Fanuc KAREL source: KT00657.KL

PROGRAM KT00657
%NOLOCKGROUP
VAR
  P1: POSITION
  P2: POSITION
  OUT: BOOLEAN
BEGIN
  OUT = + P1
END KT00657
